FUNCTION_BLOCK "FB_Motor"
{ S7_Optimized_Access := 'TRUE' }
VERSION : 0.1
   VAR_INPUT
      Enable : Bool;
   END_VAR
   VAR_OUTPUT
      Busy : Bool;
   END_VAR
BEGIN
	#Busy := #Enable AND "di_MotorFeedback";
END_FUNCTION_BLOCK
